// TIA Portal V20 export
DATA_BLOCK "CONTROL_LINE_DB"   // DB27
// stored: AutoNumber false, InstanceOfName CONTROL_LINE, InstanceOfType FB
"CONTROL_LINE"
   // VAR
   //    TIMER_reset { S7_SetPoint := 'True'} : TON_TIME;
   //    P_TRIG_INICIAL : Bool;
   //    P_TRIG_RESET : Bool;
   //    AUTOMAT { S7_SetPoint := 'True'} : "SENSOR";
   //    MANUAL { S7_SetPoint := 'True'} : "SENSOR";
   //    SENSOR_3 { S7_SetPoint := 'True'} : "SENSOR";
   //    SENSOR_4 { S7_SetPoint := 'True'} : "SENSOR";
   //    SENSOR_5 { S7_SetPoint := 'True'} : "SENSOR";
   //    SENSOR_6 { S7_SetPoint := 'True'} : "SENSOR";
   //    SENSOR_7 { S7_SetPoint := 'True'} : "SENSOR";
   //    SENSOR_8 { S7_SetPoint := 'True'} : "SENSOR";
   //    SENSOR_9 { S7_SetPoint := 'True'} : "SENSOR";
   //    SENSOR_10 { S7_SetPoint := 'True'} : "SENSOR";
   //    SENSOR_11 { S7_SetPoint := 'True'} : "SENSOR";
   //    dvere_L_A { S7_SetPoint := 'True'} : "SENSOR";
   //    dvere_L_B { S7_SetPoint := 'True'} : "SENSOR";
   //    dvere_P_A { S7_SetPoint := 'True'} : "SENSOR";
   //    dvere_P_B { S7_SetPoint := 'True'} : "SENSOR";
   //    SEN_STRUCT : Struct
   //       AUTOMAT : Bool;
   //       AUTOMAT_NEG : Bool;
   //       MANUAL : Bool;
   //       MANUAL_NEG : Bool;
   //       SENSOR_TLAKU : Bool;
   //       SENSOR_TLAKU_NEG : Bool;
   //       power : Bool;
   //       power_neg : Bool;
   //       safety : Bool;
   //       safety_neg : Bool;
   //       s_10 : Bool;
   //       TLA_STOP : Bool;
   //       TLA_STOP_NEG : Bool;
   //       TLA_START : Bool;
   //       TLA_START_NEG : Bool;
   //       TLA_KVIT : Bool;
   //       TLA_KVIT_NEG : Bool;
   //       s_17 : Bool;
   //       S19 : Bool;
   //       L1_OK : Bool;
   //       L1_NOT_OK : Bool;
   //       L2_OK : Bool;
   //       L2_NOT_OK : Bool;
   //       L3_OK : Bool;
   //       L3_NOT_OK : Bool;
   //       dvere_L_A : Bool;
   //       dvere_L_B : Bool;
   //       dvere_P_A : Bool;
   //       dvere_P_B : Bool;
   //       S30 : Bool;
   //       S31 : Bool;
   //       LASER_MEMOR : Bool;
   //    END_STRUCT;
   //    "M" : Struct
   //       P_TRIK_hmi_manual : Bool;
   //       p_trig_hmi_automat : Bool;
   //       N_TRIG_REZIM : Bool;
   //       M_4 : Bool;
   //       hlaseni_chyby : Bool;
   //       M_6 : Bool;
   //       M_7 : Bool;
   //       M_8 : Bool;
   //       M_9 : Bool;
   //       p_Trig_al : Bool;
   //       n_trig_al : Bool;
   //       p_trig_wro : Bool;
   //       n_trig_wro : Bool;
   //       M_14 : Bool;
   //       M_15 : Bool;
   //       N_TRIG_MANUAL : Bool;
   //       M_17 : Bool;
   //       M_18 : Bool;
   //       M_19 : Bool;
   //       M_20 : Bool;
   //       M_21 : Bool;
   //       M_22 : Bool;
   //       M_23 : Bool;
   //       M_24 : Bool;
   //       M_25 : Bool;
   //       M_26 : Bool;
   //       M_27 : Bool;
   //       M_28 : Bool;
   //       M_29 : Bool;
   //       M_30 : Bool;
   //       M_31 : Bool;
   //       M_32 : Bool;
   //    END_STRUCT;
   //    trig : Struct
   //       reset_error_all : Bool;
   //       TRIG_FOR_OP_4_AUTOMAT : Bool;
   //       t_3 : Bool;
   //       t_4 : Bool;
   //       t_5 : Bool;
   //       t_6 : Bool;
   //       t_7 : Bool;
   //       t_8 : Bool;
   //    END_STRUCT;
   //    SQCR : Int;
   //    job_mailbox : Array[0..3] of Word;
   //    n_trig_res_auit : Bool;
   //    inicial_control { S7_SetPoint := 'True'} : TON_TIME;
   //    SQCR_SAFETY { S7_SetPoint := 'True'} : Int;
   //    n_trig_RESET_AUT : Bool;
   //    P_TRIG_RESET_SAFETY : Bool;
   //    air { S7_SetPoint := 'True'} : TON_TIME;
   //    HMI_ALARM { S7_SetPoint := 'True'} : Int;
   // END_VAR
BEGIN
END_DATA_BLOCK
